// TIA Portal V21 export
// export: Created 2026-11-08T21:17:29.7080951Z, ExportSetting WithDefaults, DisplayName Totally Integrated Automation Portal, DisplayVersion V21 Update 3, DisplayName STEP 7 Professional, DisplayVersion V21 Update 3, DisplayName STEP 7 Safety, DisplayVersion V21, DisplayName Tech WebApplication, DisplayVersion V21, DisplayName WinCC Basic/Comfort/Advanced, DisplayVersion V21 Update 3, DisplayName WinCC Unified, DisplayVersion V21 Update 3
DATA_BLOCK "FB_Multi_DB"   // DB10
VERSION : 0.1
// stored: AutoNumber true, DBAccessibleFromOPCUA true, DBAccessibleFromWebserver true, InstanceOfName FB_Multi, InstanceOfType FB
"FB_Multi"
   // VAR_INPUT
   //    start : Bool;
   //    cfg : "UDT_Inner";
   //    mat : Array[0..1, 0..1] of Int;
   // END_VAR
   // VAR_OUTPUT
   //    done : Bool;
   // END_VAR
   // VAR_IN_OUT
   //    io : Real;
   // END_VAR
   // VAR
   //    tmr { S7_SetPoint := 'True'} : TON_TIME;
   //    tmrs { S7_SetPoint := 'True'} : Array[0..2] of TON_TIME;
   //    ctr { S7_SetPoint := 'True'} : CTU_INT;
   //    edge { S7_SetPoint := 'True'} : R_TRIG;
   //    sub { S7_SetPoint := 'True'} : "FB_Iface";
   //    subs { S7_SetPoint := 'True'} : Array[0..1] of "FB_Iface";
   //    data { S7_SetPoint := 'True'} : "UDT_Outer";
   //    cnt : Int := 8;
   //    Temp : Int;
   // END_VAR
BEGIN
   cfg.Temp := 30.0;
   mat[1,1] := 11;
   tmrs[2].PT := T#3S;
   sub.stInt := 77;
   subs[1].stInt := 78;
   data.innerArr[1].Arr[2] := 5;
END_DATA_BLOCK
